ABB RAPID module: Wobj_Wfeli.mod

MODULE Wobj_Wfeli
	! Points are read in order of declaration.
  ! Please do not change the order of points!

  LOCAL PERS robtarget pWobj_O_PointX1:=[[584.3452,-241.7878,124.3624],[0.284793198108673,-0.116733551025391,-0.951014399528503,0.0289453528821468],[-1,-1,-1,0],[9E+09,9E+09,9E+09,9E+09,9E+09,9E+09]];
	LOCAL PERS robtarget pWobj_O_PointX2:=[[410.7472,-244.4554,124.9533],[0.180527746677399,-0.264597058296204,-0.940191566944122,-0.115922264754772],[-1,-1,0,1],[9E+09,9E+09,9E+09,9E+09,9E+09,9E+09]];
	LOCAL PERS robtarget pWobj_O_PointY1:=[[588.6882,29.83716,127.4072],[0.132458090782166,0.0273857414722443,-0.989157915115356,-0.057197067886591],[0,-1,0,1],[9E+09,9E+09,9E+09,9E+09,9E+09,9E+09]];

ENDMODULE
